FUNCTION_BLOCK TcoMessengerContextTest EXTENDS TcoCore._internals_TcoContext
VAR
	_callMyPlcInstanceRtcUpdate	:	BOOL := FALSE;
	_callMyPlcInstanceRun		:	BOOL := FALSE;
	_nowLocal					:	DATE_AND_TIME;
	_nowUtc						:	DATE_AND_TIME;
	_rtcIsValid					:	BOOL := FALSE;
	_rtcIsSynchronized			:	BOOL := FALSE;
	{attribute addProperty Name "this is the name of messenger test"}
	_tcoMessangerTests			:	TcoMessengerTests(THIS^);
END_VAR

IF THIS^._callMyPlcInstanceRtcUpdate THEN
	THIS^._rtcUpdate();
	_nowLocal			:=	THIS^.RealTimeClock.NowLocal();
	_nowUtc				:=	THIS^.RealTimeClock.NowUTC();
	_rtcIsValid			:=	THIS^.RealTimeClock.IsValid;
	_rtcIsSynchronized	:=	THIS^.RealTimeClock.IsSynchronized;
END_IF

IF THIS^._callMyPlcInstanceRun THEN
	THIS^.Run();
END_IF

{attribute 'TcRpcEnable'}
METHOD INTERNAL ContextClose
SUPER^._Close();
END_METHOD

{attribute 'TcRpcEnable'}
METHOD INTERNAL ContextOpen
SUPER^._Open();
END_METHOD

METHOD PROTECTED  Main
END_METHOD

{attribute 'TcRpcEnable'}
METHOD INTERNAL RtcIsValid : BOOL
RtcIsValid := THIS^.RealTimeClock.IsValid;
_rtcIsValid := THIS^.RealTimeClock.IsValid;
END_METHOD

END_FUNCTION_BLOCK

(* stored: Version 1.1.0.1
   POU TcoMessengerContextTest: Id {ab1f1c15-693e-0b9d-1dc8-8f3fbcb09dcf}, SpecialFunc None
   Method ContextClose: Id {4f2fdfc4-fcab-0528-13d7-8604dcba8327}
   Method ContextOpen: Id {89a806dd-7d63-036b-0493-cf31446222af}
   Method Main: Id {ce1913c5-df6b-0aa3-3f90-ae6b899c0533}
   Method RtcIsValid: Id {26119aec-f827-0ffc-3e54-5571e4e4da19} *)
